Staubli VAL3: io.pjx

--- io.pjx ---
Parameters version=s8.15.3Cs9_BS3337 stackSize=5000 millimeterUnit=true
Program file=start.pgx
Program file=stop.pgx
Data file=io.dtx

--- io.dtx ---
mdesc mNomSpeed
public dio dInput[64]
public dio dOutput[64]
public aio aInput[16]
public aio aOutput[16]

--- start.pgx ---
program start()
begin
end

--- stop.pgx ---
program stop()
begin
end
